(* PLC project probe.project, CODESYS CODESYS V3.5 SP17 Patch 3 *)
(* stored: creationDateTime 2026-10-20T03:54:26.809173, modificationDateTime 1601-01-01T03:00:00 *)

FUNCTION_BLOCK FB_ProbeCfc
  VAR_INPUT
    rIn : REAL;
    rLo : REAL;
    rHi : REAL;
  END_VAR
  VAR_OUTPUT
    rOut : REAL;
  END_VAR
  VAR  (* added by the conversion: wires and edge detectors of the diagram *)
    _LIMIT1_OUT : ANY;
  END_VAR

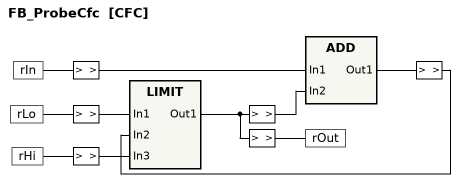
(* CFC diagram, written out as Structured Text *)
_LIMIT1_OUT := LIMIT(rLo, rIn + _LIMIT1_OUT, rHi);
rOut := _LIMIT1_OUT;
END_FUNCTION_BLOCK
